FUNCTION_BLOCK NextFeedHorizonPlant (* Basic Function Block Type *)
  (* Standard: 61499-2 *)
  (* Version 0.0, 10/19/2026, Schneider Electric, Template *)
  PACKAGE SE.Nereda;
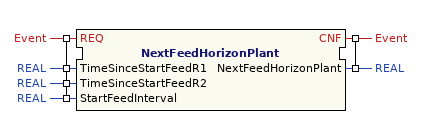
  EVENT_INPUT
    REQ WITH TimeSinceStartFeedR1, TimeSinceStartFeedR2, StartFeedInterval; (* Normal Execution Request *)
  END_EVENT
  EVENT_OUTPUT
    CNF WITH NextFeedHorizonPlant; (* Execution Confirmation *)
  END_EVENT
  VAR_INPUT
    TimeSinceStartFeedR1 : REAL;
    TimeSinceStartFeedR2 : REAL;
    StartFeedInterval : REAL;
  END_VAR
  VAR_OUTPUT
    NextFeedHorizonPlant : REAL; (* Output event qualifier *)
  END_VAR
  VAR
    LowestTimeSinceStartFeed : REAL;
  END_VAR
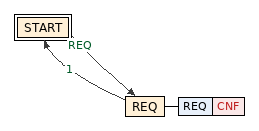
  EC_STATES
    START; (* Initial State *)
    REQ : REQ -> CNF; (* Normal execution *)
  END_STATES
  EC_TRANSITIONS
    START TO REQ := REQ;
    REQ TO START := 1;
  END_TRANSITIONS
  ALGORITHM REQ IN ST: (* Normally executed algorithm *)
;
LowestTimeSinceStartFeed := TimeSinceStartFeedR1;

IF LowestTimeSinceStartFeed > TimeSinceStartFeedR2 THEN
	LowestTimeSinceStartFeed := TimeSinceStartFeedR2;
END_IF;

NextFeedHorizonPlant := StartFeedInterval - LowestTimeSinceStartFeed;
  END_ALGORITHM
END_FUNCTION_BLOCK
